       IF #Lampentest THEN
           IF #Blink_Takt THEN #led_val:=5; ELSE #led_val:=0; END_IF;
           FOR #i:=0 TO 7 DO
               "FB_KP8_DB_1".KP8.LED[#i]:=#led_val; "FB_KP8_DB_2".KP8.LED[#i]:=#led_val; "FB_KP8_DB_3".KP8.LED[#i]:=#led_val; "FB_KP8_DB_4".KP8.LED[#i]:=#led_val;
               "FB_KP8_DB_5".KP8.LED[#i]:=#led_val; "FB_KP8_DB_6".KP8.LED[#i]:=#led_val; "FB_KP8_DB_7".KP8.LED[#i]:=#led_val; "FB_KP8_DB_8".KP8.LED[#i]:=#led_val;
               "FB_KP8_DB_9".KP8.LED[#i]:=#led_val; "FB_KP8_DB_10".KP8.LED[#i]:=#led_val; "FB_KP8_DB_11".KP8.LED[#i]:=#led_val; "FB_KP8_DB_12".KP8.LED[#i]:=#led_val;
               "FB_KP8_DB_13".KP8.LED[#i]:=#led_val; "FB_KP8_DB_14".KP8.LED[#i]:=#led_val; "FB_KP8_DB_15".KP8.LED[#i]:=#led_val; "FB_KP8_DB_16".KP8.LED[#i]:=#led_val;
               "FB_KP8_DB_17".KP8.LED[#i]:=#led_val; "FB_KP8_DB_18".KP8.LED[#i]:=#led_val; "FB_KP8_DB_19".KP8.LED[#i]:=#led_val; "FB_KP8_DB_20".KP8.LED[#i]:=#led_val;
               "FB_KP8_DB_21".KP8.LED[#i]:=#led_val; "FB_KP8_DB_22".KP8.LED[#i]:=#led_val; "FB_KP8_DB_23".KP8.LED[#i]:=#led_val; "FB_KP8_DB_24".KP8.LED[#i]:=#led_val;
               "FB_KP8_DB_25".KP8.LED[#i]:=#led_val; "FB_KP8_DB_26".KP8.LED[#i]:=#led_val; "FB_KP8_DB_27".KP8.LED[#i]:=#led_val; "FB_KP8_DB_28".KP8.LED[#i]:=#led_val;
           END_FOR;
           RETURN;
       END_IF;
       IF "DB_Bad_Konfig".Bad_Konfig[1].Hand_Aktiv_Intern THEN FOR #i:=0 TO 7 DO "FB_KP8_DB_1".KP8.LED[#i]:=3; END_FOR; END_IF;
       IF "DB_Bad_Konfig".Bad_Konfig[3].Hand_Aktiv_Intern THEN FOR #i:=0 TO 7 DO "FB_KP8_DB_2".KP8.LED[#i]:=3; END_FOR; END_IF;
       IF "DB_Bad_Konfig".Bad_Konfig[7].Hand_Aktiv_Intern THEN FOR #i:=0 TO 7 DO "FB_KP8_DB_4".KP8.LED[#i]:=3; END_FOR; END_IF;
       IF "DB_Bad_Konfig".Bad_Konfig[8].Hand_Aktiv_Intern THEN FOR #i:=0 TO 7 DO "FB_KP8_DB_5".KP8.LED[#i]:=3; END_FOR; END_IF;
       IF "DB_Bad_Konfig".Bad_Konfig[12].Hand_Aktiv_Intern THEN FOR #i:=0 TO 7 DO "FB_KP8_DB_7".KP8.LED[#i]:=3; END_FOR; END_IF;
       IF "DB_Bad_Konfig".Bad_Konfig[13].Hand_Aktiv_Intern THEN FOR #i:=0 TO 7 DO "FB_KP8_DB_8".KP8.LED[#i]:=3; END_FOR; END_IF;
       IF "DB_Bad_Konfig".Bad_Konfig[14].Hand_Aktiv_Intern THEN FOR #i:=0 TO 7 DO "FB_KP8_DB_9".KP8.LED[#i]:=3; END_FOR; END_IF;
       IF "DB_Bad_Konfig".Bad_Konfig[18].Hand_Aktiv_Intern THEN FOR #i:=0 TO 7 DO "FB_KP8_DB_11".KP8.LED[#i]:=3; END_FOR; END_IF;
       IF "DB_Bad_Konfig".Bad_Konfig[19].Hand_Aktiv_Intern THEN FOR #i:=0 TO 7 DO "FB_KP8_DB_12".KP8.LED[#i]:=3; END_FOR; END_IF;
       IF "DB_Bad_Konfig".Bad_Konfig[21].Hand_Aktiv_Intern THEN FOR #i:=0 TO 7 DO "FB_KP8_DB_13".KP8.LED[#i]:=3; END_FOR; END_IF;
       IF "DB_Bad_Konfig".Bad_Konfig[25].Hand_Aktiv_Intern THEN FOR #i:=0 TO 7 DO "FB_KP8_DB_28".KP8.LED[#i]:=3; END_FOR; END_IF;
       IF "DB_Bad_Konfig".Bad_Konfig[26].Hand_Aktiv_Intern THEN FOR #i:=0 TO 7 DO "FB_KP8_DB_15".KP8.LED[#i]:=3; END_FOR; END_IF;
       IF "DB_Bad_Konfig".Bad_Konfig[30].Hand_Aktiv_Intern THEN FOR #i:=0 TO 7 DO "FB_KP8_DB_17".KP8.LED[#i]:=3; END_FOR; END_IF;
       IF "DB_Bad_Konfig".Bad_Konfig[31].Hand_Aktiv_Intern THEN FOR #i:=0 TO 7 DO "FB_KP8_DB_18".KP8.LED[#i]:=3; END_FOR; END_IF;
       IF "DB_Bad_Konfig".Bad_Konfig[35].Hand_Aktiv_Intern THEN FOR #i:=0 TO 7 DO "FB_KP8_DB_20".KP8.LED[#i]:=3; END_FOR; END_IF;
       IF "DB_Bad_Konfig".Bad_Konfig[36].Hand_Aktiv_Intern THEN FOR #i:=0 TO 7 DO "FB_KP8_DB_21".KP8.LED[#i]:=3; END_FOR; END_IF;
       IF "DB_Bad_Konfig".Bad_Konfig[40].Hand_Aktiv_Intern THEN FOR #i:=0 TO 7 DO "FB_KP8_DB_23".KP8.LED[#i]:=3; END_FOR; END_IF;
       IF "DB_Bad_Konfig".Bad_Konfig[41].Hand_Aktiv_Intern THEN FOR #i:=0 TO 7 DO "FB_KP8_DB_24".KP8.LED[#i]:=3; END_FOR; END_IF;
       IF "DB_Bad_Konfig".Bad_Konfig[45].Hand_Aktiv_Intern THEN FOR #i:=0 TO 7 DO "FB_KP8_DB_26".KP8.LED[#i]:=3; END_FOR; END_IF;
       IF "DB_Bad_Konfig".Bad_Konfig[46].Hand_Aktiv_Intern THEN FOR #i:=0 TO 7 DO "FB_KP8_DB_27".KP8.LED[#i]:=3; END_FOR; END_IF;
       IF "DB_Bad_Konfig".Bad_Konfig[4].Hand_Aktiv_Intern OR "DB_Bad_Konfig".Bad_Konfig[5].Hand_Aktiv_Intern OR "DB_Bad_Konfig".Bad_Konfig[6].Hand_Aktiv_Intern THEN FOR #i:=0 TO 7 DO "FB_KP8_DB_3".KP8.LED[#i]:=3; END_FOR; END_IF;
       IF "DB_Bad_Konfig".Bad_Konfig[9].Hand_Aktiv_Intern OR "DB_Bad_Konfig".Bad_Konfig[10].Hand_Aktiv_Intern OR "DB_Bad_Konfig".Bad_Konfig[11].Hand_Aktiv_Intern THEN FOR #i:=0 TO 7 DO "FB_KP8_DB_6".KP8.LED[#i]:=3; END_FOR; END_IF;
       IF "DB_Bad_Konfig".Bad_Konfig[15].Hand_Aktiv_Intern OR "DB_Bad_Konfig".Bad_Konfig[16].Hand_Aktiv_Intern OR "DB_Bad_Konfig".Bad_Konfig[17].Hand_Aktiv_Intern THEN FOR #i:=0 TO 7 DO "FB_KP8_DB_10".KP8.LED[#i]:=3; END_FOR; END_IF;
       IF "DB_Bad_Konfig".Bad_Konfig[22].Hand_Aktiv_Intern OR "DB_Bad_Konfig".Bad_Konfig[23].Hand_Aktiv_Intern OR "DB_Bad_Konfig".Bad_Konfig[24].Hand_Aktiv_Intern THEN FOR #i:=0 TO 7 DO "FB_KP8_DB_14".KP8.LED[#i]:=3; END_FOR; END_IF;
       IF "DB_Bad_Konfig".Bad_Konfig[27].Hand_Aktiv_Intern OR "DB_Bad_Konfig".Bad_Konfig[28].Hand_Aktiv_Intern OR "DB_Bad_Konfig".Bad_Konfig[29].Hand_Aktiv_Intern THEN FOR #i:=0 TO 7 DO "FB_KP8_DB_16".KP8.LED[#i]:=3; END_FOR; END_IF;
       IF "DB_Bad_Konfig".Bad_Konfig[32].Hand_Aktiv_Intern OR "DB_Bad_Konfig".Bad_Konfig[33].Hand_Aktiv_Intern OR "DB_Bad_Konfig".Bad_Konfig[34].Hand_Aktiv_Intern THEN FOR #i:=0 TO 7 DO "FB_KP8_DB_19".KP8.LED[#i]:=3; END_FOR; END_IF;
       IF "DB_Bad_Konfig".Bad_Konfig[37].Hand_Aktiv_Intern OR "DB_Bad_Konfig".Bad_Konfig[38].Hand_Aktiv_Intern OR "DB_Bad_Konfig".Bad_Konfig[39].Hand_Aktiv_Intern THEN FOR #i:=0 TO 7 DO "FB_KP8_DB_22".KP8.LED[#i]:=3; END_FOR; END_IF;
       IF "DB_Bad_Konfig".Bad_Konfig[42].Hand_Aktiv_Intern OR "DB_Bad_Konfig".Bad_Konfig[43].Hand_Aktiv_Intern OR "DB_Bad_Konfig".Bad_Konfig[44].Hand_Aktiv_Intern THEN FOR #i:=0 TO 7 DO "FB_KP8_DB_25".KP8.LED[#i]:=3; END_FOR; END_IF;
END_FUNCTION

FUNCTION "FC_Not_Halt" : Void   // FC1, SCL
{ S7_Optimized_Access := 'TRUE' }
VERSION : 0.2
// stored: AutoNumber true, IsIECCheckEnabled false, SetENOAutomatically false, UDAEnableTagReadback false
   VAR_INPUT
      Not_Halt : Bool;
   END_VAR
BEGIN

       IF NOT #Not_Halt THEN RETURN; END_IF;
       "Pumpe Bad 8":=FALSE; "Pumpe Bad 12":=FALSE; "Pumpe Bad 14":=FALSE;
       "Pumpe Bad 18":=FALSE; "Pumpe Bad 19":=FALSE; "Pumpe Bad 21":=FALSE;
       "Netzschuetz Pumpe Bad 25":=FALSE;
       "FU Pumpe Freigabe":=FALSE; "Reset FU Pumpe":=FALSE;
       "Pumpen_FU_Steuerwert":=W#16#0;
       "Pumpe Bad 26":=FALSE; "Pumpe Bad 31":=FALSE; "Pumpe Bad 41":=FALSE; "Pumpe Bad 45":=FALSE;
       "Regelung Heizung Bad 7":=FALSE; "Sicherheitsschuetz Heizung Bad 7":=FALSE;
       "Regelung Heizung Bad 8":=FALSE; "Sicherheitsschuetz Heizung Bad 8":=FALSE;
       "Regelung Heizung Bad 12":=FALSE; "Sicherheitsschuetz Heizung Bad 12":=FALSE;
       "Regelung Heizung 1 Bad 25":=FALSE; "Regelung Heizung 2 Bad 25":=FALSE;
       "Sicherheitsschuetze Heizung 1 + 2 Bad 25":=FALSE;
       "Regelung Heizung Bad 36":=FALSE; "Sicherheitsschuetz Heizung Bad 36":=FALSE;
       "Regelung Heizung Bad 40":=FALSE; "Sicherheitsschuetz Heizung Bad 40":=FALSE;
       "Regelung Heizung Bad 46":=FALSE; "Sicherheitsschuetz Heizung Bad 46":=FALSE;
       "Freigabe Ultraschall Pos. 8":=FALSE; "Freigabe Ultraschall Pos. 12":=FALSE;
       "Warenbewegung 1 Bad 25 Freigabe FU":=FALSE; "Warenbewegung 1 Bad 25 Netzschuetz":=FALSE;
       "Warenbewegung 2 Bad 25 Freigabe FU":=FALSE; "Warenbewegung 2 Bad 25 Netzschuetz":=FALSE;
       "Warenbewegung 1 Bad 25 Sollwert FU":=W#16#0; "Warenbewegung 2 Bad 25 Sollwert FU":=W#16#0;
       "Masch.Leuchte 1 Anlage Hupe":=FALSE;
END_FUNCTION

FUNCTION "FC_Rueckmeldung" : Void   // FC2, SCL
{ S7_Optimized_Access := 'TRUE' }
VERSION : 0.2
// stored: AutoNumber true, IsIECCheckEnabled false, SetENOAutomatically false, UDAEnableTagReadback false
   VAR_INPUT
      Not_Halt_Aktiv : Bool;
   END_VAR
   VAR_TEMP
      "b" : Int;
      w : Int;
      ai : Int;
      si : Int;
   END_VAR
BEGIN

       "DB_CPU_to_IPC".Not_Halt_Aktiv := #Not_Halt_Aktiv;
       "DB_CPU_to_IPC".Not_Aus_OK := "Not-Aus ist OK";
       FOR #b:=1 TO "c_Anzahl_Bad" DO
           "DB_CPU_to_IPC".Bad[#b].Ampel_Status := "DB_Bad_Konfig".Bad_Konfig[#b].Ampel_Status;
           "DB_CPU_to_IPC".Bad[#b].Betriebsbereit := "DB_Bad_Konfig".Bad_Konfig[#b].Betriebsbereit;
           "DB_CPU_to_IPC".Bad[#b].Heizung_1_Ist := "DB_Bad_Konfig".Bad_Konfig[#b].Heizung_1_Ist;
           "DB_CPU_to_IPC".Bad[#b].Heizung_1_Soll := "DB_Bad_Konfig".Bad_Konfig[#b].Heizung_1_Soll;
           "DB_CPU_to_IPC".Bad[#b].Heizung_2_Ist := "DB_Bad_Konfig".Bad_Konfig[#b].Heizung_2_Ist;
           "DB_CPU_to_IPC".Bad[#b].Heizung_2_Soll := "DB_Bad_Konfig".Bad_Konfig[#b].Heizung_2_Soll;
           "DB_CPU_to_IPC".Bad[#b].Pumpe_Laeuft := "DB_Bad_Konfig".Bad_Konfig[#b].IO_Aus.Pumpe;
           "DB_CPU_to_IPC".Bad[#b].Pumpe_FU_Soll := "DB_Bad_Konfig".Bad_Konfig[#b].Pumpe_FU_Soll;
           "DB_CPU_to_IPC".Bad[#b].US_Laeuft := "DB_Bad_Konfig".Bad_Konfig[#b].IO_Aus.Ultraschall_Freigabe;
           "DB_CPU_to_IPC".Bad[#b].GR_Aktiv := "DB_Bad_Konfig".Bad_Konfig[#b].GR_Aktiv;
           "DB_CPU_to_IPC".Bad[#b].GR_Strom_Ist := "DB_Bad_Konfig".Bad_Konfig[#b].GR_Strom_Ist;
           "DB_CPU_to_IPC".Bad[#b].GR_Spannung_Ist := "DB_Bad_Konfig".Bad_Konfig[#b].GR_Spannung_Ist;
           "DB_CPU_to_IPC".Bad[#b].WB_X_Soll := "DB_Bad_Konfig".Bad_Konfig[#b].Warenbewegung_X_Soll;
           "DB_CPU_to_IPC".Bad[#b].WB_Y_Soll := "DB_Bad_Konfig".Bad_Konfig[#b].Warenbewegung_Y_Soll;
           "DB_CPU_to_IPC".Bad[#b].Hand_Aktiv := "DB_Bad_Konfig".Bad_Konfig[#b].Hand_Aktiv_Intern;
           "DB_CPU_to_IPC".Bad[#b].Hand_Abgelehnt := "DB_IPC_to_CPU".Handbetrieb[#b].Hand_Aktiv
               AND ("DB_Bad_Konfig".Bad_Konfig[#b].WT[1].Belegt OR "DB_Bad_Konfig".Bad_Konfig[#b].WT[2].Belegt OR "DB_Bad_Konfig".Bad_Konfig[#b].WT[3].Belegt);
           FOR #w:=1 TO 3 DO
               "DB_CPU_to_IPC".Bad[#b].WT[#w].Belegt := "DB_Bad_Konfig".Bad_Konfig[#b].WT[#w].Belegt;
               #ai := "DB_Bad_Konfig".Bad_Konfig[#b].WT[#w].Auftragsindex; #si := "DB_Bad_Konfig".Bad_Konfig[#b].WT[#w].SchrittIndex;
               "DB_CPU_to_IPC".Bad[#b].WT[#w].Auftragsindex := #ai; "DB_CPU_to_IPC".Bad[#b].WT[#w].SchrittIndex := #si;
               IF (#ai>=0)AND(#ai<=9)AND(#si>=0)AND(#si<=50) THEN
                   "DB_CPU_to_IPC".Bad[#b].WT[#w].Artikel_ID := "DB_IPC_to_CPU".Auftrag[#ai].ID_Artikel;
                   "DB_CPU_to_IPC".Bad[#b].WT[#w].Personal_ID := "DB_IPC_to_CPU".Auftrag[#ai].Personal_ID;
                   "DB_CPU_to_IPC".Bad[#b].WT[#w].BadNr := "DB_IPC_to_CPU".Auftrag[#ai].Schritte[#si].BadNr;
                   "DB_CPU_to_IPC".Bad[#b].WT[#w].Verweilzeit_Soll := "DB_IPC_to_CPU".Auftrag[#ai].Schritte[#si].Verweilzeit;
               END_IF;
               "DB_CPU_to_IPC".Bad[#b].WT[#w].WT_Eingesetzt := "DB_Bad_Konfig".Bad_Konfig[#b].WT[#w].WT_Eingesetzt;
               "DB_CPU_to_IPC".Bad[#b].WT[#w].Istzeit := "DB_Bad_Konfig".Bad_Konfig[#b].WT[#w].Istzeit;
               "DB_CPU_to_IPC".Bad[#b].WT[#w].Restzeit := "DB_Bad_Konfig".Bad_Konfig[#b].WT[#w].Restzeit;
               "DB_CPU_to_IPC".Bad[#b].WT[#w].Vorwarn_Erreicht := "DB_Bad_Konfig".Bad_Konfig[#b].WT[#w].Vorwarn_Erreicht;
               "DB_CPU_to_IPC".Bad[#b].WT[#w].Zeit_Abgelaufen := "DB_Bad_Konfig".Bad_Konfig[#b].WT[#w].Zeit_Abgelaufen;
               "DB_CPU_to_IPC".Bad[#b].WT[#w].Krit_Zeit_Abgelaufen := "DB_Bad_Konfig".Bad_Konfig[#b].WT[#w].Krit_Zeit_Abgelaufen;
               "DB_CPU_to_IPC".Bad[#b].WT[#w].Stoerung_Aufgetreten := "DB_Bad_Konfig".Bad_Konfig[#b].WT[#w].Stoerung_Aufgetreten;
               "DB_CPU_to_IPC".Bad[#b].WT[#w].Temp_Abweichung_Max := "DB_Bad_Konfig".Bad_Konfig[#b].WT[#w].Temp_Abweichung_Max;
               "DB_CPU_to_IPC".Bad[#b].WT[#w].Temp_Toleranz_Eingehalten := "DB_Bad_Konfig".Bad_Konfig[#b].WT[#w].Temp_Toleranz_Eingehalten;
               "DB_CPU_to_IPC".Bad[#b].WT[#w].Zeitueberschreitung := "DB_Bad_Konfig".Bad_Konfig[#b].WT[#w].Zeitueberschreitung;
               "DB_CPU_to_IPC".Bad[#b].WT[#w].Zeitstempel_Eingesetzt := "DB_Bad_Konfig".Bad_Konfig[#b].WT[#w].Zeitstempel_Eingesetzt;
               "DB_CPU_to_IPC".Bad[#b].WT[#w].Zeitstempel_Entnommen := "DB_Bad_Konfig".Bad_Konfig[#b].WT[#w].Zeitstempel_Entnommen;
               "DB_CPU_to_IPC".Bad[#b].WT[#w].Protokoll_Neu := "DB_Bad_Konfig".Bad_Konfig[#b].WT[#w].Protokoll_Neu;
           END_FOR;
       END_FOR;
END_FUNCTION

DATA_BLOCK "FB_Anlagensteuerung_DB"   // DB1
VERSION : 0.9
// stored: AutoNumber true, DBAccessibleFromOPCUA true, DBAccessibleFromWebserver true, InstanceOfName FB_Anlagensteuerung, InstanceOfType FB
"FB_Anlagensteuerung"
BEGIN
END_DATA_BLOCK

DATA_BLOCK "FB_Auftragsmanager_DB"   // DB11
VERSION : 0.1
// stored: AutoNumber true, DBAccessibleFromOPCUA true, DBAccessibleFromWebserver true, InstanceOfName FB_Auftragsmanager, InstanceOfType FB
"FB_Auftragsmanager"
BEGIN
END_DATA_BLOCK

DATA_BLOCK "FB_Bad_DB"   // DB41
VERSION : 0.2
// stored: AutoNumber true, DBAccessibleFromOPCUA true, DBAccessibleFromWebserver true, InstanceOfName FB_Bad, InstanceOfType FB
"FB_Bad"
BEGIN
END_DATA_BLOCK

DATA_BLOCK "FB_FlexKraft_DB"   // DB6
VERSION : 0.1
// stored: AutoNumber true, DBAccessibleFromOPCUA true, DBAccessibleFromWebserver true, InstanceOfName FB_FlexKraft, InstanceOfType FB
"FB_FlexKraft"
BEGIN
END_DATA_BLOCK

DATA_BLOCK "FB_FlexKraft_DB_1"   // DB7
VERSION : 0.1
// stored: AutoNumber true, DBAccessibleFromOPCUA true, DBAccessibleFromWebserver true, InstanceOfName FB_FlexKraft, InstanceOfType FB
"FB_FlexKraft"
BEGIN
END_DATA_BLOCK

DATA_BLOCK "FB_FlexKraft_DB_2"   // DB10
VERSION : 0.1
// stored: AutoNumber true, DBAccessibleFromOPCUA true, DBAccessibleFromWebserver true, InstanceOfName FB_FlexKraft, InstanceOfType FB
"FB_FlexKraft"
BEGIN
END_DATA_BLOCK

DATA_BLOCK "FB_KP8_DB_1"   // DB9
VERSION : 0.1
// stored: AutoNumber true, DBAccessibleFromOPCUA true, DBAccessibleFromWebserver true, InstanceOfName FB_Ansteuerung_KP8, InstanceOfType FB
"FB_Ansteuerung_KP8"
BEGIN
   KP8.LED[0..7] := 0;
END_DATA_BLOCK

DATA_BLOCK "FB_KP8_DB_10"   // DB20
VERSION : 0.1
// stored: AutoNumber true, DBAccessibleFromOPCUA true, DBAccessibleFromWebserver true, InstanceOfName FB_Ansteuerung_KP8, InstanceOfType FB
"FB_Ansteuerung_KP8"
BEGIN
END_DATA_BLOCK

DATA_BLOCK "FB_KP8_DB_11"   // DB21
VERSION : 0.1
// stored: AutoNumber true, DBAccessibleFromOPCUA true, DBAccessibleFromWebserver true, InstanceOfName FB_Ansteuerung_KP8, InstanceOfType FB
"FB_Ansteuerung_KP8"
BEGIN
END_DATA_BLOCK

DATA_BLOCK "FB_KP8_DB_12"   // DB22
VERSION : 0.1
// stored: AutoNumber true, DBAccessibleFromOPCUA true, DBAccessibleFromWebserver true, InstanceOfName FB_Ansteuerung_KP8, InstanceOfType FB
"FB_Ansteuerung_KP8"
BEGIN
END_DATA_BLOCK

DATA_BLOCK "FB_KP8_DB_13"   // DB23
VERSION : 0.1
// stored: AutoNumber true, DBAccessibleFromOPCUA true, DBAccessibleFromWebserver true, InstanceOfName FB_Ansteuerung_KP8, InstanceOfType FB
"FB_Ansteuerung_KP8"
BEGIN
END_DATA_BLOCK

DATA_BLOCK "FB_KP8_DB_14"   // DB24
VERSION : 0.1
// stored: AutoNumber true, DBAccessibleFromOPCUA true, DBAccessibleFromWebserver true, InstanceOfName FB_Ansteuerung_KP8, InstanceOfType FB
"FB_Ansteuerung_KP8"
BEGIN
END_DATA_BLOCK

DATA_BLOCK "FB_KP8_DB_15"   // DB25
VERSION : 0.1
// stored: AutoNumber true, DBAccessibleFromOPCUA true, DBAccessibleFromWebserver true, InstanceOfName FB_Ansteuerung_KP8, InstanceOfType FB
"FB_Ansteuerung_KP8"
BEGIN
END_DATA_BLOCK

DATA_BLOCK "FB_KP8_DB_16"   // DB26
VERSION : 0.1
// stored: AutoNumber true, DBAccessibleFromOPCUA true, DBAccessibleFromWebserver true, InstanceOfName FB_Ansteuerung_KP8, InstanceOfType FB
"FB_Ansteuerung_KP8"
BEGIN
END_DATA_BLOCK

DATA_BLOCK "FB_KP8_DB_17"   // DB27
VERSION : 0.1
// stored: AutoNumber true, DBAccessibleFromOPCUA true, DBAccessibleFromWebserver true, InstanceOfName FB_Ansteuerung_KP8, InstanceOfType FB
"FB_Ansteuerung_KP8"
BEGIN
END_DATA_BLOCK

DATA_BLOCK "FB_KP8_DB_18"   // DB28
VERSION : 0.1
// stored: AutoNumber true, DBAccessibleFromOPCUA true, DBAccessibleFromWebserver true, InstanceOfName FB_Ansteuerung_KP8, InstanceOfType FB
"FB_Ansteuerung_KP8"
BEGIN
END_DATA_BLOCK

DATA_BLOCK "FB_KP8_DB_19"   // DB29
VERSION : 0.1
// stored: AutoNumber true, DBAccessibleFromOPCUA true, DBAccessibleFromWebserver true, InstanceOfName FB_Ansteuerung_KP8, InstanceOfType FB
"FB_Ansteuerung_KP8"
BEGIN
END_DATA_BLOCK

DATA_BLOCK "FB_KP8_DB_2"   // DB12
VERSION : 0.1
// stored: AutoNumber true, DBAccessibleFromOPCUA true, DBAccessibleFromWebserver true, InstanceOfName FB_Ansteuerung_KP8, InstanceOfType FB
"FB_Ansteuerung_KP8"
BEGIN
END_DATA_BLOCK

DATA_BLOCK "FB_KP8_DB_20"   // DB30
VERSION : 0.1
// stored: AutoNumber true, DBAccessibleFromOPCUA true, DBAccessibleFromWebserver true, InstanceOfName FB_Ansteuerung_KP8, InstanceOfType FB
"FB_Ansteuerung_KP8"
BEGIN
END_DATA_BLOCK

DATA_BLOCK "FB_KP8_DB_21"   // DB31
VERSION : 0.1
// stored: AutoNumber true, DBAccessibleFromOPCUA true, DBAccessibleFromWebserver true, InstanceOfName FB_Ansteuerung_KP8, InstanceOfType FB
"FB_Ansteuerung_KP8"
BEGIN
END_DATA_BLOCK

DATA_BLOCK "FB_KP8_DB_22"   // DB32
VERSION : 0.1
// stored: AutoNumber true, DBAccessibleFromOPCUA true, DBAccessibleFromWebserver true, InstanceOfName FB_Ansteuerung_KP8, InstanceOfType FB
"FB_Ansteuerung_KP8"
BEGIN
END_DATA_BLOCK

DATA_BLOCK "FB_KP8_DB_23"   // DB33
VERSION : 0.1
// stored: AutoNumber true, DBAccessibleFromOPCUA true, DBAccessibleFromWebserver true, InstanceOfName FB_Ansteuerung_KP8, InstanceOfType FB
"FB_Ansteuerung_KP8"
BEGIN
END_DATA_BLOCK

DATA_BLOCK "FB_KP8_DB_24"   // DB34
VERSION : 0.1
// stored: AutoNumber true, DBAccessibleFromOPCUA true, DBAccessibleFromWebserver true, InstanceOfName FB_Ansteuerung_KP8, InstanceOfType FB
"FB_Ansteuerung_KP8"
BEGIN
END_DATA_BLOCK

DATA_BLOCK "FB_KP8_DB_25"   // DB35
VERSION : 0.1
// stored: AutoNumber true, DBAccessibleFromOPCUA true, DBAccessibleFromWebserver true, InstanceOfName FB_Ansteuerung_KP8, InstanceOfType FB
"FB_Ansteuerung_KP8"
BEGIN
END_DATA_BLOCK

DATA_BLOCK "FB_KP8_DB_26"   // DB36
VERSION : 0.1
// stored: AutoNumber true, DBAccessibleFromOPCUA true, DBAccessibleFromWebserver true, InstanceOfName FB_Ansteuerung_KP8, InstanceOfType FB
"FB_Ansteuerung_KP8"
BEGIN
END_DATA_BLOCK

DATA_BLOCK "FB_KP8_DB_27"   // DB37
VERSION : 0.1
// stored: AutoNumber true, DBAccessibleFromOPCUA true, DBAccessibleFromWebserver true, InstanceOfName FB_Ansteuerung_KP8, InstanceOfType FB
"FB_Ansteuerung_KP8"
BEGIN
END_DATA_BLOCK

DATA_BLOCK "FB_KP8_DB_28"   // DB38
VERSION : 0.1
// stored: AutoNumber true, DBAccessibleFromOPCUA true, DBAccessibleFromWebserver true, InstanceOfName FB_Ansteuerung_KP8, InstanceOfType FB
"FB_Ansteuerung_KP8"
BEGIN
END_DATA_BLOCK

DATA_BLOCK "FB_KP8_DB_3"   // DB13
VERSION : 0.1
// stored: AutoNumber true, DBAccessibleFromOPCUA true, DBAccessibleFromWebserver true, InstanceOfName FB_Ansteuerung_KP8, InstanceOfType FB
"FB_Ansteuerung_KP8"
BEGIN
END_DATA_BLOCK

DATA_BLOCK "FB_KP8_DB_4"   // DB14
VERSION : 0.1
// stored: AutoNumber true, DBAccessibleFromOPCUA true, DBAccessibleFromWebserver true, InstanceOfName FB_Ansteuerung_KP8, InstanceOfType FB
"FB_Ansteuerung_KP8"
BEGIN
END_DATA_BLOCK

DATA_BLOCK "FB_KP8_DB_5"   // DB15
VERSION : 0.1
// stored: AutoNumber true, DBAccessibleFromOPCUA true, DBAccessibleFromWebserver true, InstanceOfName FB_Ansteuerung_KP8, InstanceOfType FB
"FB_Ansteuerung_KP8"
BEGIN
END_DATA_BLOCK

DATA_BLOCK "FB_KP8_DB_6"   // DB16
VERSION : 0.1
// stored: AutoNumber true, DBAccessibleFromOPCUA true, DBAccessibleFromWebserver true, InstanceOfName FB_Ansteuerung_KP8, InstanceOfType FB
"FB_Ansteuerung_KP8"
BEGIN
END_DATA_BLOCK

DATA_BLOCK "FB_KP8_DB_7"   // DB17
VERSION : 0.1
// stored: AutoNumber true, DBAccessibleFromOPCUA true, DBAccessibleFromWebserver true, InstanceOfName FB_Ansteuerung_KP8, InstanceOfType FB
"FB_Ansteuerung_KP8"
BEGIN
END_DATA_BLOCK

DATA_BLOCK "FB_KP8_DB_8"   // DB18
VERSION : 0.1
// stored: AutoNumber true, DBAccessibleFromOPCUA true, DBAccessibleFromWebserver true, InstanceOfName FB_Ansteuerung_KP8, InstanceOfType FB
"FB_Ansteuerung_KP8"
BEGIN
END_DATA_BLOCK

DATA_BLOCK "FB_KP8_DB_9"   // DB19
VERSION : 0.1
// stored: AutoNumber true, DBAccessibleFromOPCUA true, DBAccessibleFromWebserver true, InstanceOfName FB_Ansteuerung_KP8, InstanceOfType FB
"FB_Ansteuerung_KP8"
BEGIN
END_DATA_BLOCK
